FUNCTION_BLOCK NextFeedHorizonCalc2 (* Basic Function Block Type *)
  (* Standard: 61499-2 *)
  (* Version 0.0, 7/15/2026, Schneider Electric, Template *)
  PACKAGE SE.Nereda;
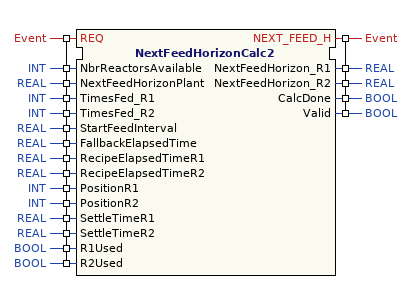
  EVENT_INPUT
    REQ WITH StartFeedInterval, PositionR1, PositionR2, SettleTimeR1, SettleTimeR2, FallbackElapsedTime, R1Used, R2Used, TimesFed_R1, TimesFed_R2, NbrReactorsAvailable, RecipeElapsedTimeR1, RecipeElapsedTimeR2, NextFeedHorizonPlant;
  END_EVENT
  EVENT_OUTPUT
    NEXT_FEED_H WITH NextFeedHorizon_R2, NextFeedHorizon_R1, CalcDone, Valid;
  END_EVENT
  VAR_INPUT
    NbrReactorsAvailable : INT;
    NextFeedHorizonPlant : REAL;
    TimesFed_R1 : INT; (* = 0 the First Feed *)
    TimesFed_R2 : INT;
    StartFeedInterval : REAL;
    FallbackElapsedTime : REAL;
    RecipeElapsedTimeR1 : REAL;
    RecipeElapsedTimeR2 : REAL;
    PositionR1 : INT;
    PositionR2 : INT;
    SettleTimeR1 : REAL;
    SettleTimeR2 : REAL;
    R1Used : BOOL;
    R2Used : BOOL;
  END_VAR
  VAR_OUTPUT
    NextFeedHorizon_R1 : REAL;
    NextFeedHorizon_R2 : REAL;
    CalcDone : BOOL;
    Valid : BOOL;
  END_VAR
  VAR
    InNextFeedHorizon_R1 : REAL;
    InNextFeedHorizon_R2 : REAL;
    InNextFeedHorizon_R3 : REAL;
    InNextFeedHorizon_R4 : REAL;
    InNextFeedHorizon_R5 : REAL;
    InNextFeedHorizon_R6 : REAL;
  END_VAR
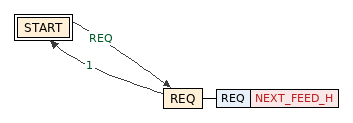
  EC_STATES
    START; (* Initial State *)
    REQ : REQ -> NEXT_FEED_H; (* Normal execution *)
  END_STATES
  EC_TRANSITIONS
    START TO REQ := REQ;
    REQ TO START := 1;
  END_TRANSITIONS
  ALGORITHM REQ IN ST: (* Normally executed algorithm *)
// Validation
Valid := (FallbackElapsedTime > 0) AND (StartFeedInterval > 0);

// Calculate Next Feed Horizon for each Reactor
IF Valid THEN
	IF R1Used THEN
		IF TimesFed_R1 = 0 THEN
			InNextFeedHorizon_R1 := (PositionR1 - 1) * StartFeedInterval - FallbackElapsedTime + SettleTimeR1;
		ELSE
			//InNextFeedHorizon_R1 := (NbrReactorsAvailable * StartFeedInterval) - RecipeElapsedTimeR1;
			InNextFeedHorizon_R1 := NextFeedHorizonPlant + (StartFeedInterval * (PositionR1 - 1));
		END_IF;
	END_IF;

	IF R2Used THEN
		IF TimesFed_R2 = 0 THEN
			InNextFeedHorizon_R2 := (PositionR2 - 1) * StartFeedInterval - FallbackElapsedTime + SettleTimeR2;
		ELSE
			//InNextFeedHorizon_R2 := (NbrReactorsAvailable * StartFeedInterval) - RecipeElapsedTimeR2;
			InNextFeedHorizon_R2 := NextFeedHorizonPlant + (StartFeedInterval * (PositionR2 - 1));
		END_IF;
	END_IF;
END_IF;

//Verify Calculation
CalcDone := Valid AND (InNextFeedHorizon_R1 <> 0 OR InNextFeedHorizon_R2 <> 0);

//Results
IF InNextFeedHorizon_R1 > 0 THEN
    NextFeedHorizon_R1 := InNextFeedHorizon_R1;
ELSE
    NextFeedHorizon_R1 := 0;
END_IF;

IF InNextFeedHorizon_R2 > 0 THEN
    NextFeedHorizon_R2 := InNextFeedHorizon_R2;
ELSE
    NextFeedHorizon_R2 := 0;
END_IF;
  END_ALGORITHM
END_FUNCTION_BLOCK
